// TIA Portal V20 export
VAR_GLOBAL   // PLC tag table "Default tag table"
   RESERVE_AI_1 AT %IW66 : Int;
   "System_Byte(1)" AT %MB1 : Byte;
   reset_hsc AT %M2.7 : Bool;
END_VAR
